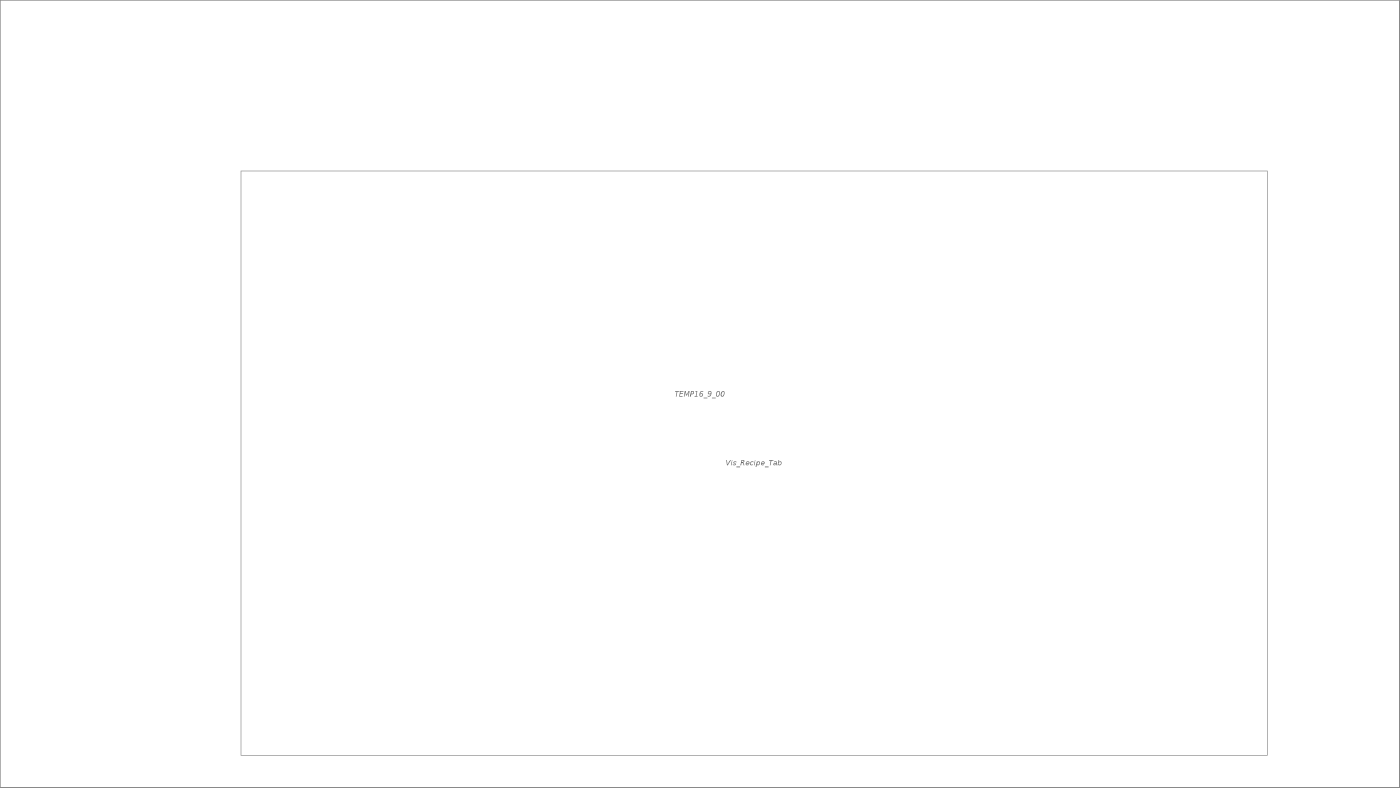
VISUALIZATION Recipe_16_9  // 1920x1081
    Frame (0,0 1920x1081)
        shows TEMP16_9_00()
    Frame (330,234 1408x802)
        shows Vis_Recipe_Tab()
END_VISUALIZATION

(* stored: Version 1.1.0.1, ProductVersion 3.1.4024.13
   Visu Recipe_16_9: Id {00ce2abd-1f96-44eb-ad0d-6adabb5160fa} *)
